FUNCTION_BLOCK F (* Positive: two waiting positions, exits on an input *)
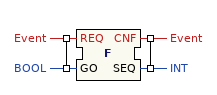
  EVENT_INPUT
    REQ WITH GO;
  END_EVENT
  EVENT_OUTPUT
    CNF WITH SEQ;
  END_EVENT
  VAR_INPUT
    GO : BOOL;
  END_VAR
  VAR_OUTPUT
    SEQ : INT;
  END_VAR
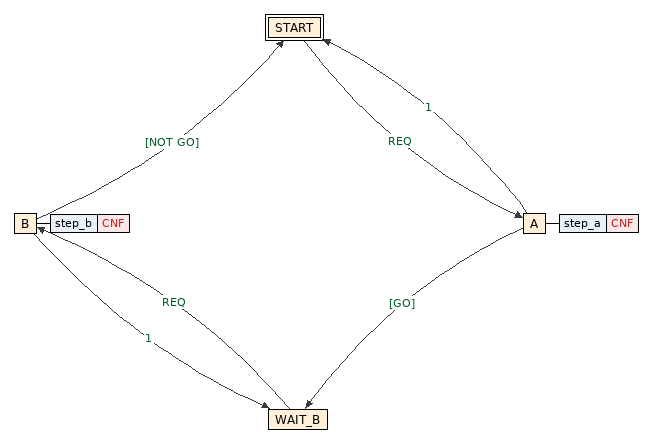
  EC_STATES
    START;
    A : step_a -> CNF;
    WAIT_B;
    B : step_b -> CNF;
  END_STATES
  EC_TRANSITIONS
    START TO A := REQ;
    A TO WAIT_B := [GO];
    A TO START := 1;
    WAIT_B TO B := REQ;
    B TO START := [NOT GO];
    B TO WAIT_B := 1;
  END_TRANSITIONS
  ALGORITHM step_a IN ST:
SEQ := 0;
IF GO THEN
  SEQ := 1;
END_IF;
  END_ALGORITHM
  ALGORITHM step_b IN ST:
IF NOT GO THEN
  SEQ := 0;
END_IF;
  END_ALGORITHM
END_FUNCTION_BLOCK
